(* IEC 61131-3 sources: nautilus/examples/pump-station, 3 files *)

(* ---- motor.st ---- *)
(* A root .st file with no PROGRAM is a library: it is in scope for every
   task's compile, so `type: Motor` in the manifest resolves against it.
   On an EtherNet/IP project you do not write this file — `nautilus eip
   import` emits eip_types.st from the controller's own UDT definitions. *)

TYPE
  Motor : STRUCT
    Running : BOOL;
    Fault   : BOOL;
    Speed   : REAL;
    Hours   : REAL;
  END_STRUCT;
END_TYPE

(* ---- sim.st ---- *)
PROGRAM Sim
(* Stands in for the field bus: writes the Motor structs that a real
   deployment's EtherNet/IP driver would supply.

   NOTE THE SHAPE. `P101.Running := ...` on a VAR_EXTERNAL struct compiles
   and runs (the VM read-modify-writes the tag). This file keeps the older
   form — copy → mutate the LOCAL → assign the whole struct back — because
   it rewrites most of the struct each scan, and that is one tag write
   instead of a dozen. Either form is correct. *)
VAR_EXTERNAL
    P101 : Motor;  P101_Enable : BOOL;  P101_StartSP : REAL;
    P102 : Motor;  P102_Enable : BOOL;  P102_StartSP : REAL;
    P103 : Motor;  P103_Enable : BOOL;  P103_StartSP : REAL;
    P201 : Motor;  P201_Enable : BOOL;  P201_StartSP : REAL;
    P202 : Motor;  P202_Enable : BOOL;  P202_StartSP : REAL;
    P301 : Motor;  P301_Enable : BOOL;  P301_StartSP : REAL;
END_VAR
VAR
    m : Motor;
END_VAR

m := P101; m.Running := P101_Enable AND NOT m.Fault;
IF m.Running THEN m.Speed := P101_StartSP; ELSE m.Speed := 0.0; END_IF; P101 := m;

m := P102; m.Running := P102_Enable AND NOT m.Fault;
IF m.Running THEN m.Speed := P102_StartSP; ELSE m.Speed := 0.0; END_IF; P102 := m;

m := P103; m.Running := P103_Enable AND NOT m.Fault;
IF m.Running THEN m.Speed := P103_StartSP; ELSE m.Speed := 0.0; END_IF; P103 := m;

m := P201; m.Running := P201_Enable AND NOT m.Fault;
IF m.Running THEN m.Speed := P201_StartSP; ELSE m.Speed := 0.0; END_IF; P201 := m;

m := P202; m.Running := P202_Enable AND NOT m.Fault;
IF m.Running THEN m.Speed := P202_StartSP; ELSE m.Speed := 0.0; END_IF; P202 := m;

m := P301; m.Running := P301_Enable AND NOT m.Fault;
IF m.Running THEN m.Speed := P301_StartSP; ELSE m.Speed := 0.0; END_IF; P301 := m;

END_PROGRAM

(* ---- station.st ---- *)
PROGRAM Station
(* Per-pump logic. This is the part the design brief is honest about NOT
   shortening: the manifest holds 24 tags from 9 authored rows, but the
   VAR_EXTERNAL block below is still one line per tag. `nautilus eip import`
   emits a ready-to-paste block for exactly this reason. *)
VAR_EXTERNAL
    P101 : Motor;  P101_RunHrs : REAL;  P101_StartSP : REAL;  P101_Enable : BOOL;
    P102 : Motor;  P102_RunHrs : REAL;  P102_StartSP : REAL;  P102_Enable : BOOL;
    P103 : Motor;  P103_RunHrs : REAL;  P103_StartSP : REAL;  P103_Enable : BOOL;
    P201 : Motor;  P201_RunHrs : REAL;  P201_StartSP : REAL;  P201_Enable : BOOL;
    P202 : Motor;  P202_RunHrs : REAL;  P202_StartSP : REAL;  P202_Enable : BOOL;
    P301 : Motor;  P301_RunHrs : REAL;  P301_StartSP : REAL;  P301_Enable : BOOL;
    StationDtS  : REAL;
    RunningCount : REAL;
    AnyFault     : BOOL;
END_VAR

(* run-hour accumulation, per pump *)
IF P101.Running THEN P101_RunHrs := P101_RunHrs + StationDtS / 3600.0; END_IF;
IF P102.Running THEN P102_RunHrs := P102_RunHrs + StationDtS / 3600.0; END_IF;
IF P103.Running THEN P103_RunHrs := P103_RunHrs + StationDtS / 3600.0; END_IF;
IF P201.Running THEN P201_RunHrs := P201_RunHrs + StationDtS / 3600.0; END_IF;
IF P202.Running THEN P202_RunHrs := P202_RunHrs + StationDtS / 3600.0; END_IF;
IF P301.Running THEN P301_RunHrs := P301_RunHrs + StationDtS / 3600.0; END_IF;

(* station rollups — the tags an operator screen actually shows *)
RunningCount := 0.0;
IF P101.Running THEN RunningCount := RunningCount + 1.0; END_IF;
IF P102.Running THEN RunningCount := RunningCount + 1.0; END_IF;
IF P103.Running THEN RunningCount := RunningCount + 1.0; END_IF;
IF P201.Running THEN RunningCount := RunningCount + 1.0; END_IF;
IF P202.Running THEN RunningCount := RunningCount + 1.0; END_IF;
IF P301.Running THEN RunningCount := RunningCount + 1.0; END_IF;

AnyFault := P101.Fault OR P102.Fault OR P103.Fault
         OR P201.Fault OR P202.Fault OR P301.Fault;

END_PROGRAM
